PROGRAM Branches
  VAR
    w01_a : BOOL;
    w01_y : BOOL;
    w01_b : BOOL;
    w01_e : BOOL;
    w01_c : BOOL;
    w01_d : BOOL;
    w02_f : BOOL;
    w02_y : BOOL;
    w02_g : BOOL;
    w02_j : BOOL;
    w02_h : BOOL;
    w02_i : BOOL;
    w02_k : BOOL;
    w03_e : BOOL;
    w03_y : BOOL;
    w03_a : BOOL;
    w03_b : BOOL;
    w03_d : BOOL;
    w03_c : BOOL;
    w04_a : BOOL;
    w04_y : BOOL;
    w04_conveyor_infeed_photoeye_blocked_longer_than_limit : BOOL;
    w04_b : BOOL;
    w05_a : BOOL;
    w05_k : BOOL;
    w05_conveyor_reject_gate_solenoid_output_main : BOOL;
  END_VAR

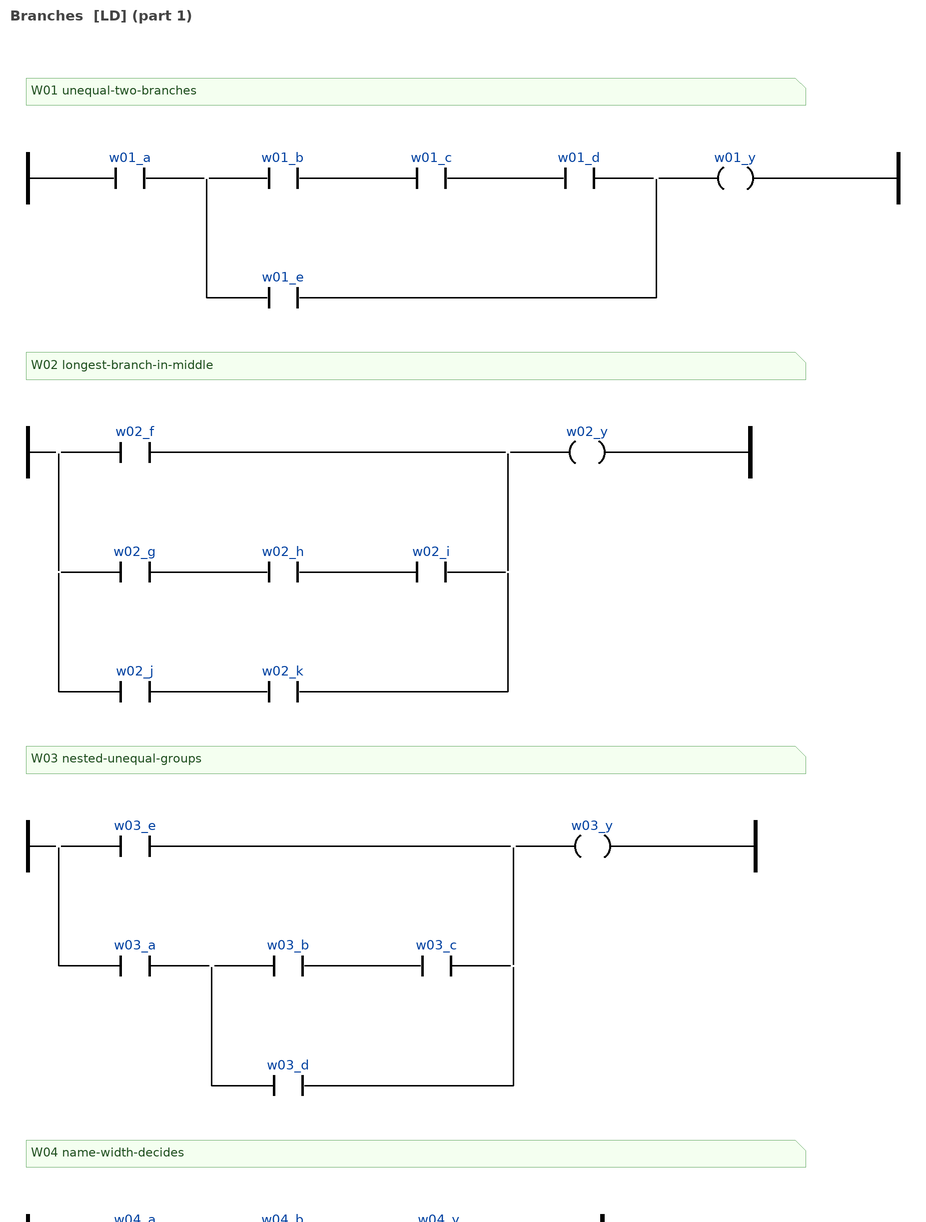
(* LD diagram, written out as Structured Text *)
(* W01 unequal-two-branches *)
w01_y := w01_a AND (w01_e OR w01_b AND w01_c AND w01_d);
(* W02 longest-branch-in-middle *)
w02_y := w02_f OR w02_g AND w02_h AND w02_i OR w02_j AND w02_k;
(* W03 nested-unequal-groups *)
w03_y := w03_e OR w03_a AND w03_d OR w03_a AND w03_b AND w03_c;
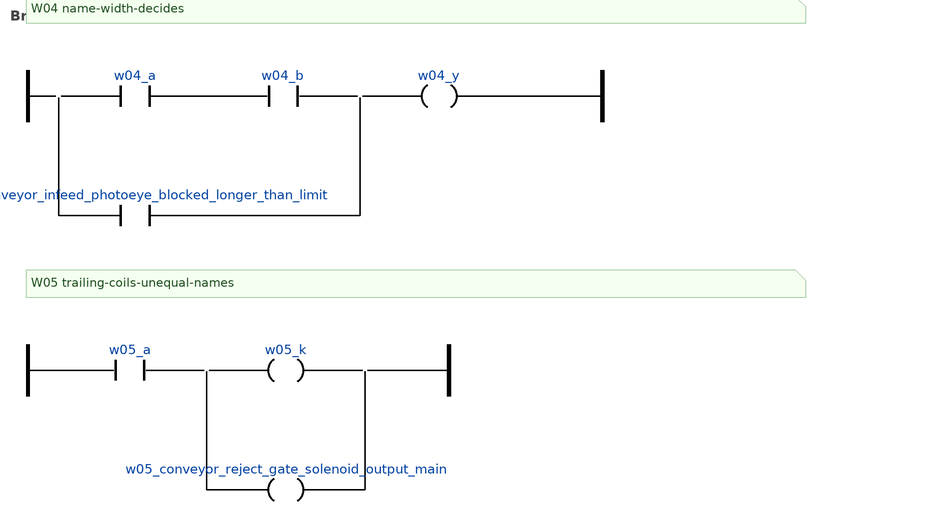
(* W04 name-width-decides *)
w04_y := w04_conveyor_infeed_photoeye_blocked_longer_than_limit OR w04_a AND w04_b;
(* W05 trailing-coils-unequal-names *)
w05_k := w05_a;
w05_conveyor_reject_gate_solenoid_output_main := w05_a;
END_PROGRAM
